(* IEC 61131-3 sources: plc-st-coding-agent/progress/evidence/full_r8_20261110b/native_evidence/codex_minimax-m27/self-hard-05/1, 1 file *)

(* ---- candidate.st ---- *)
FUNCTION_BLOCK FB
VAR_INPUT
    runRequest  : BOOL;
    flameOK     : BOOL;
    o2Valid     : BOOL;
    o2PV        : REAL;
    baseAir     : REAL;
    resetBtn    : BOOL;
END_VAR
VAR_OUTPUT
    fuelPermit  : BOOL;
    trimEnable  : BOOL;
    airTrim     : REAL;
    airCommand  : REAL;
    tripLatched : BOOL;
    o2Fault     : BOOL;
END_VAR
VAR
    prevResetBtn : BOOL := FALSE;
    resetRising  : BOOL;
END_VAR

resetRising := resetBtn AND NOT prevResetBtn;

IF runRequest AND NOT flameOK THEN
    tripLatched := TRUE;
ELSIF resetRising AND NOT runRequest AND NOT flameOK THEN
    tripLatched := FALSE;
END_IF

prevResetBtn := resetBtn;

fuelPermit := runRequest AND flameOK AND NOT tripLatched;

o2Fault := NOT o2Valid OR o2PV < 0.0 OR o2PV > 21.0;

trimEnable := fuelPermit AND NOT o2Fault;

IF trimEnable THEN
    airTrim := 2.0 * (2.0 - o2PV);
    IF airTrim > 10.0 THEN
        airTrim := 10.0;
    ELSIF airTrim < -10.0 THEN
        airTrim := -10.0;
    END_IF
ELSE
    airTrim := 0.0;
END_IF

IF fuelPermit THEN
    airCommand := baseAir + airTrim;
    IF airCommand > 100.0 THEN
        airCommand := 100.0;
    ELSIF airCommand < 0.0 THEN
        airCommand := 0.0;
    END_IF
ELSE
    airCommand := 0.0;
END_IF

END_FUNCTION_BLOCK
